TYPE "ST_PressDemoParCfg"
VERSION : 0.1
   STRUCT
      SchemaVersion : UInt := 3;
      IdealCycleMs : UDInt := 0;
      BaselineWorkMs : UDInt := 0;
      Timeout : Time := T#10S;
      TransferSettleTime : Time := T#100MS;
      PressSettleTime : Time := T#500MS;
   END_STRUCT;

END_TYPE

